(* IEC 61131-3 sources: s7-to-codesys/src/POUs/S7Compat/F_S5CountUp, 2 files *)

(* ---- F_S5CountUp.decl.st ---- *)
// Назначение: CU C n — счёт вверх счётчика S5: по фронту RLO 0 → 1 значение +1, не больше 999 (AWL_e.pdf,
//             гл. 4). Возвращает значение после инструкции.
// Автор:      kr0nsch
// Версия:     1.2.0
// Документ:   docs/MAPPING_STL.md, правило s5.counter
FUNCTION F_S5CountUp : INT
VAR_IN_OUT
    stCounter : ST_S5Counter;   // счётчик (GVL_S5Counters.aCounter[n])
END_VAR
VAR_INPUT
    xRlo : BOOL;                // RLO перед инструкцией
END_VAR
VAR CONSTANT
    MAX_VALUE : INT := 999;     // верхняя граница счётчика S5
END_VAR

(* ---- F_S5CountUp.impl.st ---- *)
IF xRlo AND NOT stCounter.xRloUp AND stCounter.iValue < MAX_VALUE THEN
    stCounter.iValue := stCounter.iValue + 1;
END_IF
stCounter.xRloUp := xRlo;
F_S5CountUp := stCounter.iValue;
